// Tests for MONETcommon.F_CommandAcceptance and F_CommandRejectText (#83, #87): one test per row of the
// acceptance table (specs/plans/2026-10-20-command-acceptance-83-87.md, section 2.2).
FUNCTION_BLOCK F_CommandAcceptance_Tests EXTENDS TcUnit.FB_TestSuite
VAR
	eLastReason	: MONETcommon.E_CommandRejectReason;
END_VAR

Ready_Idle_Accepts_All();
Estop_Rejects_Moves_Accepts_Park();
Error_Rejects_Moves_Accepts_Park();
Clock_Invalid_Rejects_All_Moves_Except_GoHome();
Stopping_Rejects_Moves_Defers_Park();
Powering_Rejects_Moves_Park_Aborts_Power();
Parking_Rejects_Moves();
Parked_Rejects_Moves_With_Reason_Parked();
Parked_Park_Is_Accepted();
InitRequired_Rejects_Moves_Accepts_Park();
NotReady_Rejects_Moves_Accepts_Park();
GoHome_Active_Rejects_Slew_Goto_Track();
Moving_Replaces();
Reject_Texts();
Reject_Reason_Maps_To_Brotlib();

// A powered-on, idle telescope: nothing pending, nothing wrong.
METHOD PRIVATE Ready_State : MONETcommon.ST_CommandState
Ready_State.bClockValid := TRUE;
Ready_State.bReady := TRUE;
END_METHOD

METHOD PRIVATE Decide : MONETcommon.E_CommandDecision
VAR_INPUT
	eCommand	: BROTLib.E_TCSCommand;
	stState		: MONETcommon.ST_CommandState;
END_VAR
Decide := MONETcommon.F_CommandAcceptance(eCommand := eCommand, stState := stState, eReason => eLastReason);
END_METHOD

METHOD PRIVATE Ready_Idle_Accepts_All
VAR
	stState	: MONETcommon.ST_CommandState;
END_VAR
TEST('Ready_Idle_Accepts_All');
stState := Ready_State();
AssertTrue(Condition := Decide(BROTLib.E_TCSCommand.slew, stState) = MONETcommon.E_CommandDecision.accept, Message := 'slew');
AssertTrue(Condition := Decide(BROTLib.E_TCSCommand.goto, stState) = MONETcommon.E_CommandDecision.accept, Message := 'goto');
AssertTrue(Condition := Decide(BROTLib.E_TCSCommand.track, stState) = MONETcommon.E_CommandDecision.accept, Message := 'track');
AssertTrue(Condition := Decide(BROTLib.E_TCSCommand.gohome, stState) = MONETcommon.E_CommandDecision.accept, Message := 'gohome');
AssertTrue(Condition := Decide(BROTLib.E_TCSCommand.park, stState) = MONETcommon.E_CommandDecision.accept, Message := 'park');
AssertTrue(Condition := eLastReason = MONETcommon.E_CommandRejectReason.none, Message := 'no reason on accept');
TEST_FINISHED();
END_METHOD

METHOD PRIVATE Estop_Rejects_Moves_Accepts_Park
VAR
	stState	: MONETcommon.ST_CommandState;
END_VAR
TEST('Estop_Rejects_Moves_Accepts_Park');
stState := Ready_State();
stState.bEstop := TRUE;
stState.bError := TRUE;		// the E-stop also raises an error: the E-stop reason wins
AssertTrue(Condition := Decide(BROTLib.E_TCSCommand.slew, stState) = MONETcommon.E_CommandDecision.reject, Message := 'slew rejected');
AssertTrue(Condition := eLastReason = MONETcommon.E_CommandRejectReason.estop, Message := 'reason estop');
AssertTrue(Condition := Decide(BROTLib.E_TCSCommand.gohome, stState) = MONETcommon.E_CommandDecision.reject, Message := 'gohome rejected');
AssertTrue(Condition := Decide(BROTLib.E_TCSCommand.park, stState) = MONETcommon.E_CommandDecision.accept, Message := 'park accepted');
TEST_FINISHED();
END_METHOD

// The emergency park (#86 is out of scope) must stay reachable: park is accepted with an error.
METHOD PRIVATE Error_Rejects_Moves_Accepts_Park
VAR
	stState	: MONETcommon.ST_CommandState;
END_VAR
TEST('Error_Rejects_Moves_Accepts_Park');
stState := Ready_State();
stState.bError := TRUE;
stState.bReady := FALSE;
stState.bIsParked := TRUE;		// error beats parked
AssertTrue(Condition := Decide(BROTLib.E_TCSCommand.goto, stState) = MONETcommon.E_CommandDecision.reject, Message := 'goto rejected');
AssertTrue(Condition := eLastReason = MONETcommon.E_CommandRejectReason.error, Message := 'reason error');
AssertTrue(Condition := Decide(BROTLib.E_TCSCommand.park, stState) = MONETcommon.E_CommandDecision.accept, Message := 'park accepted');
stState.bPowering := TRUE;		// an error during a power-on: no abort branch, the error path handles it
AssertTrue(Condition := Decide(BROTLib.E_TCSCommand.park, stState) = MONETcommon.E_CommandDecision.accept, Message := 'park accepted while powering with error');
TEST_FINISHED();
END_METHOD

METHOD PRIVATE Clock_Invalid_Rejects_All_Moves_Except_GoHome
VAR
	stState	: MONETcommon.ST_CommandState;
END_VAR
TEST('Clock_Invalid_Rejects_All_Moves_Except_GoHome');
stState := Ready_State();
stState.bClockValid := FALSE;
AssertTrue(Condition := Decide(BROTLib.E_TCSCommand.slew, stState) = MONETcommon.E_CommandDecision.reject, Message := 'slew rejected');
AssertTrue(Condition := eLastReason = MONETcommon.E_CommandRejectReason.clock_invalid, Message := 'reason clock');
AssertTrue(Condition := Decide(BROTLib.E_TCSCommand.goto, stState) = MONETcommon.E_CommandDecision.reject, Message := 'goto rejected');
AssertTrue(Condition := Decide(BROTLib.E_TCSCommand.track, stState) = MONETcommon.E_CommandDecision.reject, Message := 'track rejected');
AssertTrue(Condition := Decide(BROTLib.E_TCSCommand.gohome, stState) = MONETcommon.E_CommandDecision.accept, Message := 'gohome needs no time');
AssertTrue(Condition := Decide(BROTLib.E_TCSCommand.park, stState) = MONETcommon.E_CommandDecision.accept, Message := 'park accepted');
TEST_FINISHED();
END_METHOD

METHOD PRIVATE Stopping_Rejects_Moves_Defers_Park
VAR
	stState	: MONETcommon.ST_CommandState;
END_VAR
TEST('Stopping_Rejects_Moves_Defers_Park');
stState := Ready_State();
stState.bStop := TRUE;
stState.bPowering := TRUE;		// a stop beats a power-on
AssertTrue(Condition := Decide(BROTLib.E_TCSCommand.slew, stState) = MONETcommon.E_CommandDecision.reject, Message := 'slew rejected');
AssertTrue(Condition := eLastReason = MONETcommon.E_CommandRejectReason.stopping, Message := 'reason stopping');
AssertTrue(Condition := Decide(BROTLib.E_TCSCommand.gohome, stState) = MONETcommon.E_CommandDecision.reject, Message := 'gohome rejected');
AssertTrue(Condition := Decide(BROTLib.E_TCSCommand.park, stState) = MONETcommon.E_CommandDecision.defer, Message := 'park deferred to standstill');
TEST_FINISHED();
END_METHOD

METHOD PRIVATE Powering_Rejects_Moves_Park_Aborts_Power
VAR
	stState	: MONETcommon.ST_CommandState;
END_VAR
TEST('Powering_Rejects_Moves_Park_Aborts_Power');
stState := Ready_State();
stState.bPowering := TRUE;
stState.bReady := FALSE;
stState.bIsParked := TRUE;		// power-on starts from parked: "power-on in progress" wins over "parked"
AssertTrue(Condition := Decide(BROTLib.E_TCSCommand.goto, stState) = MONETcommon.E_CommandDecision.reject, Message := 'goto rejected');
AssertTrue(Condition := eLastReason = MONETcommon.E_CommandRejectReason.powering_on, Message := 'reason powering_on');
AssertTrue(Condition := Decide(BROTLib.E_TCSCommand.track, stState) = MONETcommon.E_CommandDecision.reject, Message := 'track rejected');
AssertTrue(Condition := Decide(BROTLib.E_TCSCommand.park, stState) = MONETcommon.E_CommandDecision.abort_power, Message := '#87 park aborts the power-on');
TEST_FINISHED();
END_METHOD

METHOD PRIVATE Parking_Rejects_Moves
VAR
	stState	: MONETcommon.ST_CommandState;
END_VAR
TEST('Parking_Rejects_Moves');
stState := Ready_State();
stState.bParkPending := TRUE;
AssertTrue(Condition := Decide(BROTLib.E_TCSCommand.slew, stState) = MONETcommon.E_CommandDecision.reject, Message := 'slew rejected');
AssertTrue(Condition := eLastReason = MONETcommon.E_CommandRejectReason.parking, Message := 'reason parking');
AssertTrue(Condition := Decide(BROTLib.E_TCSCommand.gohome, stState) = MONETcommon.E_CommandDecision.reject, Message := 'gohome rejected');
AssertTrue(Condition := Decide(BROTLib.E_TCSCommand.park, stState) = MONETcommon.E_CommandDecision.accept, Message := 'park again is a no-op accept');
TEST_FINISHED();
END_METHOD

// #83: a slew sent to a parked telescope is rejected at once and never stays pending.
METHOD PRIVATE Parked_Rejects_Moves_With_Reason_Parked
VAR
	stState	: MONETcommon.ST_CommandState;
END_VAR
TEST('Parked_Rejects_Moves_With_Reason_Parked');
stState := Ready_State();
stState.bIsParked := TRUE;
stState.bReady := FALSE;
AssertTrue(Condition := Decide(BROTLib.E_TCSCommand.slew, stState) = MONETcommon.E_CommandDecision.reject, Message := 'slew rejected');
AssertTrue(Condition := eLastReason = MONETcommon.E_CommandRejectReason.parked, Message := 'slew reason parked');
AssertTrue(Condition := Decide(BROTLib.E_TCSCommand.goto, stState) = MONETcommon.E_CommandDecision.reject, Message := 'goto rejected');
AssertTrue(Condition := Decide(BROTLib.E_TCSCommand.track, stState) = MONETcommon.E_CommandDecision.reject, Message := 'track rejected');
AssertTrue(Condition := Decide(BROTLib.E_TCSCommand.gohome, stState) = MONETcommon.E_CommandDecision.reject, Message := 'gohome rejected');
AssertTrue(Condition := eLastReason = MONETcommon.E_CommandRejectReason.parked, Message := 'gohome reason parked');
TEST_FINISHED();
END_METHOD

// #72: after manual mode every move is rejected with init_required, park stays accepted, the earlier rows keep their reason
// and a FALSE latch changes nothing.
METHOD PRIVATE InitRequired_Rejects_Moves_Accepts_Park
VAR
	stState	: MONETcommon.ST_CommandState;
END_VAR
TEST('InitRequired_Rejects_Moves_Accepts_Park');
stState := Ready_State();
stState.bInitRequired := TRUE;
AssertTrue(Condition := Decide(BROTLib.E_TCSCommand.slew, stState) = MONETcommon.E_CommandDecision.reject, Message := 'slew rejected');
AssertTrue(Condition := eLastReason = MONETcommon.E_CommandRejectReason.init_required, Message := 'reason init_required (slew)');
AssertTrue(Condition := Decide(BROTLib.E_TCSCommand.goto, stState) = MONETcommon.E_CommandDecision.reject, Message := 'goto rejected');
AssertTrue(Condition := Decide(BROTLib.E_TCSCommand.track, stState) = MONETcommon.E_CommandDecision.reject, Message := 'track rejected');
AssertTrue(Condition := Decide(BROTLib.E_TCSCommand.gohome, stState) = MONETcommon.E_CommandDecision.reject, Message := 'gohome rejected');
AssertTrue(Condition := eLastReason = MONETcommon.E_CommandRejectReason.init_required, Message := 'reason init_required (gohome)');
AssertTrue(Condition := Decide(BROTLib.E_TCSCommand.park, stState) = MONETcommon.E_CommandDecision.accept, Message := 'park accepted');
// the rows above it keep their reason
stState.bEstop := TRUE;
AssertTrue(Condition := Decide(BROTLib.E_TCSCommand.slew, stState) = MONETcommon.E_CommandDecision.reject, Message := 'estop: rejected');
AssertTrue(Condition := eLastReason = MONETcommon.E_CommandRejectReason.estop, Message := 'estop keeps precedence');
stState.bEstop := FALSE;
stState.bIsParked := TRUE;
AssertTrue(Condition := Decide(BROTLib.E_TCSCommand.slew, stState) = MONETcommon.E_CommandDecision.reject, Message := 'parked: rejected');
AssertTrue(Condition := eLastReason = MONETcommon.E_CommandRejectReason.parked, Message := 'parked keeps precedence');
// without the latch nothing changes
stState := Ready_State();
AssertTrue(Condition := Decide(BROTLib.E_TCSCommand.slew, stState) = MONETcommon.E_CommandDecision.accept, Message := 'no latch: accepted');
TEST_FINISHED();
END_METHOD

METHOD PRIVATE Parked_Park_Is_Accepted
VAR
	stState	: MONETcommon.ST_CommandState;
END_VAR
TEST('Parked_Park_Is_Accepted');
stState := Ready_State();
stState.bIsParked := TRUE;
stState.bReady := FALSE;
AssertTrue(Condition := Decide(BROTLib.E_TCSCommand.park, stState) = MONETcommon.E_CommandDecision.accept, Message := 'park accepted');
AssertTrue(Condition := eLastReason = MONETcommon.E_CommandRejectReason.none, Message := 'no reason');
TEST_FINISHED();
END_METHOD

METHOD PRIVATE NotReady_Rejects_Moves_Accepts_Park
VAR
	stState	: MONETcommon.ST_CommandState;
END_VAR
TEST('NotReady_Rejects_Moves_Accepts_Park');
stState := Ready_State();
stState.bReady := FALSE;
AssertTrue(Condition := Decide(BROTLib.E_TCSCommand.slew, stState) = MONETcommon.E_CommandDecision.reject, Message := 'slew rejected');
AssertTrue(Condition := eLastReason = MONETcommon.E_CommandRejectReason.not_ready, Message := 'reason not_ready');
AssertTrue(Condition := Decide(BROTLib.E_TCSCommand.gohome, stState) = MONETcommon.E_CommandDecision.reject, Message := 'gohome rejected');
AssertTrue(Condition := Decide(BROTLib.E_TCSCommand.park, stState) = MONETcommon.E_CommandDecision.accept, Message := 'park accepted');
TEST_FINISHED();
END_METHOD

METHOD PRIVATE GoHome_Active_Rejects_Slew_Goto_Track
VAR
	stState	: MONETcommon.ST_CommandState;
END_VAR
TEST('GoHome_Active_Rejects_Slew_Goto_Track');
stState := Ready_State();
stState.bGoHomeActive := TRUE;
stState.bMoveActive := TRUE;
AssertTrue(Condition := Decide(BROTLib.E_TCSCommand.slew, stState) = MONETcommon.E_CommandDecision.reject, Message := 'slew rejected');
AssertTrue(Condition := eLastReason = MONETcommon.E_CommandRejectReason.gohome_active, Message := 'reason gohome_active');
AssertTrue(Condition := Decide(BROTLib.E_TCSCommand.goto, stState) = MONETcommon.E_CommandDecision.reject, Message := 'goto rejected');
AssertTrue(Condition := Decide(BROTLib.E_TCSCommand.track, stState) = MONETcommon.E_CommandDecision.reject, Message := 'track rejected');
AssertTrue(Condition := Decide(BROTLib.E_TCSCommand.gohome, stState) = MONETcommon.E_CommandDecision.replace, Message := 'gohome over gohome replaces');
AssertTrue(Condition := Decide(BROTLib.E_TCSCommand.park, stState) = MONETcommon.E_CommandDecision.accept, Message := 'park accepted');
TEST_FINISHED();
END_METHOD

// Latest move wins: slew over goto, goto over slew, goto over tracking, gohome over a move.
METHOD PRIVATE Moving_Replaces
VAR
	stState	: MONETcommon.ST_CommandState;
END_VAR
TEST('Moving_Replaces');
stState := Ready_State();
stState.bMoveActive := TRUE;
AssertTrue(Condition := Decide(BROTLib.E_TCSCommand.slew, stState) = MONETcommon.E_CommandDecision.replace, Message := 'slew replaces');
AssertTrue(Condition := Decide(BROTLib.E_TCSCommand.goto, stState) = MONETcommon.E_CommandDecision.replace, Message := 'goto replaces');
AssertTrue(Condition := Decide(BROTLib.E_TCSCommand.track, stState) = MONETcommon.E_CommandDecision.replace, Message := 'track replaces');
AssertTrue(Condition := Decide(BROTLib.E_TCSCommand.gohome, stState) = MONETcommon.E_CommandDecision.replace, Message := 'gohome replaces');
AssertTrue(Condition := eLastReason = MONETcommon.E_CommandRejectReason.none, Message := 'no reason on replace');
AssertTrue(Condition := Decide(BROTLib.E_TCSCommand.park, stState) = MONETcommon.E_CommandDecision.accept, Message := 'park is not a replace');
TEST_FINISHED();
END_METHOD

// every reason except none has a log text
METHOD PRIVATE Reject_Texts
VAR
	eReason	: MONETcommon.E_CommandRejectReason;
END_VAR
TEST('Reject_Texts');
AssertEquals_STRING(Expected := '', Actual := MONETcommon.F_CommandRejectText(MONETcommon.E_CommandRejectReason.none), Message := 'none has no text');
eReason := MONETcommon.E_CommandRejectReason.estop;
AssertTrue(Condition := LEN(MONETcommon.F_CommandRejectText(eReason)) > 0, Message := 'estop');
eReason := MONETcommon.E_CommandRejectReason.error;
AssertTrue(Condition := LEN(MONETcommon.F_CommandRejectText(eReason)) > 0, Message := 'error');
eReason := MONETcommon.E_CommandRejectReason.clock_invalid;
AssertTrue(Condition := LEN(MONETcommon.F_CommandRejectText(eReason)) > 0, Message := 'clock_invalid');
eReason := MONETcommon.E_CommandRejectReason.stopping;
AssertTrue(Condition := LEN(MONETcommon.F_CommandRejectText(eReason)) > 0, Message := 'stopping');
eReason := MONETcommon.E_CommandRejectReason.powering_on;
AssertTrue(Condition := LEN(MONETcommon.F_CommandRejectText(eReason)) > 0, Message := 'powering_on');
eReason := MONETcommon.E_CommandRejectReason.parking;
AssertTrue(Condition := LEN(MONETcommon.F_CommandRejectText(eReason)) > 0, Message := 'parking');
eReason := MONETcommon.E_CommandRejectReason.parked;
AssertTrue(Condition := LEN(MONETcommon.F_CommandRejectText(eReason)) > 0, Message := 'parked');
eReason := MONETcommon.E_CommandRejectReason.not_ready;
AssertTrue(Condition := LEN(MONETcommon.F_CommandRejectText(eReason)) > 0, Message := 'not_ready');
eReason := MONETcommon.E_CommandRejectReason.gohome_active;
AssertTrue(Condition := LEN(MONETcommon.F_CommandRejectText(eReason)) > 0, Message := 'gohome_active');
eReason := MONETcommon.E_CommandRejectReason.init_required;
AssertEquals_STRING(Expected := 'init required after manual mode, send power=1 first', Actual := MONETcommon.F_CommandRejectText(eReason), Message := 'init_required text (#72)');
AssertEquals_STRING(Expected := 'telescope parked, send power=1 first', Actual := MONETcommon.F_CommandRejectText(MONETcommon.E_CommandRejectReason.parked), Message := 'parked text (#83)');
TEST_FINISHED();
END_METHOD

// X2: the local reject reason reaches I_TelescopeStatus.LastRejectReason as the BROTLib enum, member by member.
METHOD PRIVATE Reject_Reason_Maps_To_Brotlib
TEST('Reject_Reason_Maps_To_Brotlib');
AssertTrue(Condition := MONETcommon.F_RejectReasonToBrotlib(eReason := MONETcommon.E_CommandRejectReason.none) = BROTLib.E_CommandRejectReason.none, Message := 'none');
AssertTrue(Condition := MONETcommon.F_RejectReasonToBrotlib(eReason := MONETcommon.E_CommandRejectReason.estop) = BROTLib.E_CommandRejectReason.estop, Message := 'estop');
AssertTrue(Condition := MONETcommon.F_RejectReasonToBrotlib(eReason := MONETcommon.E_CommandRejectReason.error) = BROTLib.E_CommandRejectReason.error, Message := 'error');
AssertTrue(Condition := MONETcommon.F_RejectReasonToBrotlib(eReason := MONETcommon.E_CommandRejectReason.clock_invalid) = BROTLib.E_CommandRejectReason.clock_invalid, Message := 'clock_invalid');
AssertTrue(Condition := MONETcommon.F_RejectReasonToBrotlib(eReason := MONETcommon.E_CommandRejectReason.stopping) = BROTLib.E_CommandRejectReason.stopping, Message := 'stopping');
AssertTrue(Condition := MONETcommon.F_RejectReasonToBrotlib(eReason := MONETcommon.E_CommandRejectReason.powering_on) = BROTLib.E_CommandRejectReason.powering_on, Message := 'powering_on');
AssertTrue(Condition := MONETcommon.F_RejectReasonToBrotlib(eReason := MONETcommon.E_CommandRejectReason.parking) = BROTLib.E_CommandRejectReason.parking, Message := 'parking');
AssertTrue(Condition := MONETcommon.F_RejectReasonToBrotlib(eReason := MONETcommon.E_CommandRejectReason.parked) = BROTLib.E_CommandRejectReason.parked, Message := 'parked');
AssertTrue(Condition := MONETcommon.F_RejectReasonToBrotlib(eReason := MONETcommon.E_CommandRejectReason.not_ready) = BROTLib.E_CommandRejectReason.not_ready, Message := 'not_ready');
AssertTrue(Condition := MONETcommon.F_RejectReasonToBrotlib(eReason := MONETcommon.E_CommandRejectReason.gohome_active) = BROTLib.E_CommandRejectReason.gohome_active, Message := 'gohome_active');
AssertTrue(Condition := MONETcommon.F_RejectReasonToBrotlib(eReason := MONETcommon.E_CommandRejectReason.init_required) = BROTLib.E_CommandRejectReason.init_required, Message := 'init_required');
TEST_FINISHED();
END_METHOD

END_FUNCTION_BLOCK

(* stored: Version 1.1.0.1, ProductVersion 3.1.4024.15
   POU F_CommandAcceptance_Tests: Id {5b1d2a10-7c3e-4d52-9a61-0e4f8c2b7a21}, SpecialFunc None
   Method Ready_State: Id {5b1d2a10-7c3e-4d52-9a61-0e4f8c2b7a22}
   Method Decide: Id {5b1d2a10-7c3e-4d52-9a61-0e4f8c2b7a23}
   Method Ready_Idle_Accepts_All: Id {5b1d2a10-7c3e-4d52-9a61-0e4f8c2b7a24}
   Method Estop_Rejects_Moves_Accepts_Park: Id {5b1d2a10-7c3e-4d52-9a61-0e4f8c2b7a25}
   Method Error_Rejects_Moves_Accepts_Park: Id {5b1d2a10-7c3e-4d52-9a61-0e4f8c2b7a26}
   Method Clock_Invalid_Rejects_All_Moves_Except_GoHome: Id {5b1d2a10-7c3e-4d52-9a61-0e4f8c2b7a27}
   Method Stopping_Rejects_Moves_Defers_Park: Id {5b1d2a10-7c3e-4d52-9a61-0e4f8c2b7a28}
   Method Powering_Rejects_Moves_Park_Aborts_Power: Id {5b1d2a10-7c3e-4d52-9a61-0e4f8c2b7a29}
   Method Parking_Rejects_Moves: Id {5b1d2a10-7c3e-4d52-9a61-0e4f8c2b7a2a}
   Method Parked_Rejects_Moves_With_Reason_Parked: Id {5b1d2a10-7c3e-4d52-9a61-0e4f8c2b7a2b}
   Method InitRequired_Rejects_Moves_Accepts_Park: Id {72b3d6f1-8a4c-4e17-b5d9-3c0a91e7f274}
   Method Parked_Park_Is_Accepted: Id {5b1d2a10-7c3e-4d52-9a61-0e4f8c2b7a2c}
   Method NotReady_Rejects_Moves_Accepts_Park: Id {5b1d2a10-7c3e-4d52-9a61-0e4f8c2b7a2d}
   Method GoHome_Active_Rejects_Slew_Goto_Track: Id {5b1d2a10-7c3e-4d52-9a61-0e4f8c2b7a2e}
   Method Moving_Replaces: Id {5b1d2a10-7c3e-4d52-9a61-0e4f8c2b7a2f}
   Method Reject_Texts: Id {5b1d2a10-7c3e-4d52-9a61-0e4f8c2b7a30}
   Method Reject_Reason_Maps_To_Brotlib: Id {404b8666-467e-4515-97fe-dbe64c60e49e} *)
